{attribute 'Tc2GvlVarNames'}
VAR_GLOBAL
	stgGr02Alarm			:ST_AlarmRef;
END_VAR

(* stored: Version 1.1.0.1, ProductVersion 3.1.4024.15
   GVL GVL_Gr02Alarm: Id {8be4b255-3451-40e3-9f73-a18ba44fcfeb} *)
